GLOBALCONSTANTS FU_Demo_Konstanten (* Adressen der FU-Demo: Modbus-TCP-Verbindungen (APIXON -> Waveshare RS232/485/422 TO POE ETH (B) -> DELIXI H300 0,75 kW) und lokale OPC-UA-Knoten fuer das Web-Dashboard. Alle Adressen, IPs und Skalierungen nur hier aendern. *)
  (* Standard: 61499-1; Description: Copyright (c) 2026 Franz Höpfinger This program and the accompanying materials are made available under the terms of the Eclipse Public License 2.0 which is available at https://www.eclipse.org/legal/epl-2.0/ SPDX-License-Identifier: EPL-2.0 *)
  (* Version 1.1, 2026-11-02, Franz Höpfinger, Franz Höpfinger, FU_SYSTEM_TICK_WEB_WRITE (Lebenszeichen fuer das Dashboard). *)
  (* Version 1.0, 2026-11-02, Franz Höpfinger, Franz Höpfinger, initial - ein H300 an einem Waveshare-Gateway, Register laut H300-Handbuch Kap. 9.1 / 9.2.9. *)
  PACKAGE FBs::FU_Demo;
  VAR_GLOBAL CONSTANT
    APIXON : WSTRING := "192.168.1.11:61499"; (* MGR_ID der APIXON (Deploy-Adresse der 4diac IDE) - einzige Stelle *)
    FU_MODBUS_LESEN : WSTRING := "modbus[tcp:192.168.1.200:4196:1:500:h36864..36868,h36870,h37682,h37683:]"; (* Zyklisches Lesen (500 ms), Adressen DEZIMAL (FORTE parst mit strtoul Basis 10!): 36864..36868 = *)
    FU_MODBUS_KOMMANDO : WSTRING := "modbus[tcp:192.168.1.200:4196:1:500::h37632]"; (* Steuerwort 9300H = 37632 dezimal (1=Vorwaerts, 2=Rueckwaerts, 5=Freier Auslauf, 6=Rampenstopp, *)
    FU_MODBUS_SOLLWERT : WSTRING := "modbus[tcp:192.168.1.200:4196:1:500::h37633]"; (* Frequenzsollwert 9301H = 37633 dezimal, 0..10000 = 0,00..100,00 % von P0.1.16 (Maximalfrequenz), *)
    FU_FMAX_HZ : REAL := 80.0; (* Muss zu P0.1.16 (Maximalfrequenz) UND P0.1.18 (obere Grenzfrequenz) am Umrichter passen, beide am 2026-11-02 auf 80,00 Hz gesetzt *)
    FU_SOLLWERT_FAKTOR : REAL := REAL#125.0; (* Hz -> Registerwert 9301H: 10000 / FU_FMAX_HZ (125.0 bei 80 Hz) - bei Aenderung von FU_FMAX_HZ mit anpassen. Typisiertes Literal REAL#, weil es an den generischen Eingang F_MUL.IN2 geht. *)
    FU_SKALIERUNG_0_01 : REAL := 0.01; (* Registerauflösung 0,01 (Frequenz in Hz, Strom in A) *)
    FU_SKALIERUNG_0_1 : REAL := 0.1; (* Registerauflösung 0,1 (Zwischenkreisspannung in V, Leistung in kW) *)
    FU_SKALIERUNG_1 : REAL := 1.0; (* Registerauflösung 1 (Ausgangsspannung in V) *)
    FU_MESSWERTE_WEB_WRITE : WSTRING := "opc_ua[WRITE;/Objects/FU1/IstFrequenz,1:s=FU1.IstFrequenz;/Objects/FU1/SollFrequenzAktiv,1:s=FU1.SollFrequenzAktiv;/Objects/FU1/Strom,1:s=FU1.Strom;/Objects/FU1/Ausgangsspannung,1:s=FU1.Ausgangsspannung;/Objects/FU1/Zwischenkreisspannung,1:s=FU1.Zwischenkreisspannung;/Objects/FU1/Leistung,1:s=FU1.Leistung;/Objects/FU1/Status,1:s=FU1.Status;/Objects/FU1/Fehlercode,1:s=FU1.Fehlercode]"; (* PUBLISH_8 auf den lokalen OPC-UA-Server, vom Web-Dashboard abonniert. Reihenfolge = SD_1..SD_8. *)
    FU_KOMMANDO_WEB_READ : WSTRING := "opc_ua[READ;/Objects/FU1/Kommando,1:s=FU1.Kommando]"; (* Steuerwort vom Web-Dashboard (UInt16, Werte siehe FU_MODBUS_KOMMANDO). Jeder Schreibzugriff des *)
    FU_SOLLFREQUENZ_WEB_READ : WSTRING := "opc_ua[READ;/Objects/FU1/SollFrequenz,1:s=FU1.SollFrequenz]"; (* Sollfrequenz in Hz vom Web-Dashboard (Float), wird auf 0..FU_FMAX_HZ begrenzt *)
    FU_SYSTEM_TICK_WEB_WRITE : WSTRING := "opc_ua[WRITE;/Objects/FU1/System/Tick,1:s=FU1.SYSTEM_TICK]"; (* Lebenszeichen 0..99 alle 200 ms fuer das Web-Dashboard *)
  END_VAR
END_GLOBALCONSTANTS
